// TIA Portal V20 export
DATA_BLOCK "Main_Safety_RTG1_DB"   // DB15, F_DB
NAME : FUSI
// stored: InstanceOfName Main_Safety_RTG1, InstanceOfType FB
"Main_Safety_RTG1"
   // VAR
   //    "ESTOP1_NOT-HALT Taster1" : ESTOP1;
   //    "stat_Q_NOT-HALT Taster1" : Bool;
   //    "stat_AckReq_NOT-HALT Taster1" : Bool;
   //    "ESTOP1_NOT-HALT Extern 1" : ESTOP1;
   //    "stat_Q_NOT-HALT Extern 1" : Bool;
   //    "stat_AckReq_NOT-HALT Extern1" : Bool;
   //    "ESTOP1_NOT-HALT Extern 2" : ESTOP1;
   //    "stat_Q_NOT-HALT Extern 2" : Bool;
   //    "stat_AckReq_NOT-HALT Extern 2" : Bool;
   //    "ESTOP1_Tür 1" : ESTOP1;
   //    "stat_Q_Tür 1" : Bool;
   //    "stat_AckReq_Tür 1" : Bool;
   //    "ESTOP1_Tür 2" : ESTOP1;
   //    "stat_Q_Tür 2" : Bool;
   //    "stat_AckReq_Tür 2" : Bool;
   //    ESTOP1_Systemdruck : ESTOP1;
   //    stat_AckReq_Systemdruck : Bool;
   //    "FDBACK_1_NOT-HALT Schütz mit DE_NOT-HALT_Schuetz_Rueckf" : FDBACK;
   //    "stat_Q_FDBK_1_NOT-HALT Schütz mit DE_NOT-HALT_Schuetz_Rueckf" : Bool;
   //    "stat_ERROR_FDBK_1_NOT-HALT Schütz mit DE_NOT-HALT_Schuetz_Rueckf" : Bool;
   //    "FDBACK_2_NOT-HALT Schütz mit IS_Rueck_Entlueftung" : FDBACK;
   //    "stat_Q_FDBK_2_NOT-HALT Schütz mit IS_Rueck_Entlueftung" : Bool;
   //    "stat_ERROR_FDBK_2_NOT-HALT Schütz mit IS_Rueck_Entlueftung" : Bool;
   //    "FDBACK_3_NOT-HALT Schütz mit IS_Druckbereich_entlueftet" : FDBACK;
   //    "stat_Q_FDBK_3_NOT-HALT Schütz mit IS_Druckbereich_entlueftet" : Bool;
   //    "stat_ERROR_FDBK_3_NOT-HALT Schütz mit IS_Druckbereich_entlueftet" : Bool;
   //    "FDBACK_4_NOT-HALT Türe 1 RST mit DE_NOT-HALT_Tuere_1_Rueck_RST" : FDBACK;
   //    "stat_Q_FDBK_4_NOT-HALT Türe 1 RST mit DE_NOT-HALT_Tuere_1_Rueck_RST" : Bool;
   //    "stat_ERROR_FDBK_4_NOT-HALT Türe 1 RST mit DE_NOT-HALT_Tuere_1_Rueck_RST" : Bool;
   //    "FDBACK_5_NOT-HALT Türe 1 mit DE_NOT-HALT_Tuere_1_Rueckf" : FDBACK;
   //    "stat_Q_FDBK_5_NOT-HALT Türe 1 mit DE_NOT-HALT_Tuere_1_Rueckf" : Bool;
   //    "stat_ERROR_FDBK_5_NOT-HALT Türe 1 mit DE_NOT-HALT_Tuere_1_Rueckf" : Bool;
   //    "FDBACK_6_NOT-HALT Türe 1 mit DE_Antriebe_Rueckf" : FDBACK;
   //    "stat_Q_FDBK_6_NOT-HALT Türe 1 mit DE_Antriebe_Rueckf" : Bool;
   //    "stat_ERROR_FDBK_6_NOT-HALT Türe 1 mit DE_Antriebe_Rueckf" : Bool;
   //    "FDBACK_7_NOT-HALT Türe 2 RST mit DE_NOT-HALT_Tuere_2_Rueck_RST" : FDBACK;
   //    "stat_Q_FDBK_7_NOT-HALT Türe 2 RST mit DE_NOT-HALT_Tuere_2_Rueck_RST" : Bool;
   //    "stat_ERROR_FDBK_7_NOT-HALT Türe 2 RST mit DE_NOT-HALT_Tuere_2_Rueck_RST" : Bool;
   //    "FDBACK_8_NOT-HALT Türe 2 mit DE_NOT-HALT_Tuere_2_Rueckf" : FDBACK;
   //    "stat_Q_FDBK_8_NOT-HALT Türe 2 mit DE_NOT-HALT_Tuere_2_Rueckf" : Bool;
   //    "stat_ERROR_FDBK_8_NOT-HALT Türe 2 mit DE_NOT-HALT_Tuere_2_Rueckf" : Bool;
   //    "FDBACK_10_Sicherere Bewegung" : FDBACK;
   //    "stat_AckReq_10_Sicherere Bewegung" : Bool;
   //    ACK_GL_Instance : ACK_GL;
   //    Systemdruck_OK : Bool;
   //    Antriebe_sicher : Bool;
   //    "TON_Zuhaltung_Freigben_mit_NOT-HALT" : TON;
   //    BA_0_groesser_1_5 : Bool;
   //    TON_BA_0_groesser_1_5 : TON;
   //    TON_Türen_setzen_zum_öffnen : TON;
   //    BA_0 : Bool;
   //    Zuhaltung_freigegeben : Bool;
   // END_VAR
BEGIN
END_DATA_BLOCK
